(* PLC project Vn_ld_reset_coil, Beckhoff Automation GmbH TwinCAT PLC Control 3.5.13.21 *)
(* stored: creationDateTime 1970-01-01T00:00:00 *)

PROGRAM Vn_ld_reset_coil

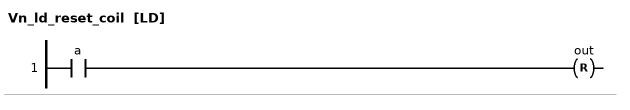
(* LD diagram, written out as Structured Text *)
IF a THEN out := FALSE; END_IF;
END_PROGRAM
